(* CODESYS project tccamera.library
   Company: TcNexa
   DefaultNamespace: TcNexa_Devices_Camera_TcCamera
   Version: 1.0.0.0
   Placeholder: TcCamera
   Author: ATI Software Engineering
   Title: TcCamera

Project tree, tasks and I/O mapping:
  libraries: Tc2_Standard, * (Beckhoff Automation GmbH); Tc2_System, * (Beckhoff Automation GmbH); Tc3_Module, * (Beckhoff Automation GmbH); TcProcess, * (TcNexa)
  ITFs/
    interface I_Camera: inRunMode, inspect, setProgramNumber
  Tests/
    program PRG_TEST [ST]
  Version/
    global variables Global_Version
*)

// Version/Global_Version
{attribute 'TcGenerated'}
{attribute 'no-analysis'}
{attribute 'linkalways'}
// This function has been automatically generated from the project information.
VAR_GLOBAL CONSTANT
	{attribute 'const_non_replaced'}
	stLibVersion_TcCamera : ST_LibVersion := (iMajor := 1, iMinor := 0, iBuild := 0, iRevision := 0, nFlags := 0, sVersion := '1.0.0.0');
END_VAR

// ITFs/I_Camera
INTERFACE I_Camera

PROPERTY inRunMode : BOOL
GET
END_GET
END_PROPERTY

METHOD inspect
VAR_INPUT
	Response		: REFERENCE TO TcNexa_Components_TcProcess.FB_MethodResponse;
END_VAR
END_METHOD

METHOD setProgramNumber
VAR_INPUT
	programNumber	: UINT;
	Response		: REFERENCE TO TcNexa_Components_TcProcess.FB_MethodResponse;
END_VAR
END_METHOD

END_INTERFACE

// Tests/PRG_TEST
PROGRAM PRG_TEST
VAR
END_VAR

END_PROGRAM
